Fanuc KAREL source: kb00112.KL

-- PROVISIONAL review KL for V770-1; original PC SHA256 5cec90b09c4bb7d454155a4b37ee17bb781d22db9f22ed52c465b4ad29963900
-- Incomplete behavior may be omitted. Consult companion uncertainty JSON. Do not deploy.
PROGRAM KB00112
%NOLOCKGROUP
VAR
  RESULT : BOOLEAN
-- UNRESOLVED_DECL P1 type=000199
BEGIN
  -- UNRESOLVED_PC offsets 5-28; opcodes 27,22,1C,27,9D,76,23
  -- UNRESOLVED_PC offsets 33-37; opcodes 7F
END KB00112
